// TIA Portal project "000_empty" (V21)

(* hardware
DEVICE "PLC_1"  S7-1500 station
   slot 0: "Rail_0"  Rack  6ES7 590-1***0-0AA0
   slot 1: "PLC_1"  CPU 1513-1 PN  6ES7 513-1AL02-0AB0  V2.9
      slot 3: "CPU display_1"  6ES7591-1AA00-0AA0
      slot 32768: "PROFINET interface_1"  X1
         slot 32769: "Port_1"  X1 P1
         slot 32770: "Port_2"  X1 P2
      slot 34817: "Virtual CP interface port_1"  Virtual CP interface port  Virtual CP interface port
*)

// ===== PLC "PLC_1"  CPU 1513-1 PN =====

VAR_GLOBAL   // PLC tag table "Default tag table"
   "Tag__639296449648259132" AT %MW10 : Word;
   "Tag__639296449652422717" AT %MW12 : Word;
   "Tag__639296449666761157" AT %T1 : Timer;
   "Tag__639296449667118790" AT %T2 : Timer;
   "Tag__639296449667279911" AT %T3 : Timer;
   "Tag__639296449667396582" AT %T4 : Timer;
   "Tag__639296449667490544" AT %T5 : Timer;
   "Tag__639296449667666479" AT %C1 : Counter;
END_VAR

TYPE "UDT_Motor"
   STRUCT
      Running : Bool;   // Motor on
      Speed : Real := 1500.0;   // Speed setpoint
      Count : Int := 7;
   END_STRUCT;
END_TYPE

DATA_BLOCK "DB_Global"   // DB1
{ S7_Optimized_Access := 'TRUE' }
   VAR
      xBool : Bool := TRUE;   // Bool comment
      iInt : Int := 42;
      rReal : Real := 3.5;   // Real comment
      aInt : Array[0..3] of Int;
      sData : Struct
         "a" : Bool;
         "b" : DInt := -5;
      END_STRUCT;
   END_VAR
BEGIN
   aInt[1] := 11;
END_DATA_BLOCK

DATA_BLOCK "FB_Empty_DB"   // DB2
{ S7_Optimized_Access := 'TRUE' }
VERSION : 0.1
// stored: InstanceOfName FB_Empty
"FB_Empty"
BEGIN
END_DATA_BLOCK

DATA_BLOCK "DB_Motor"   // DB4
{ S7_Optimized_Access := 'TRUE' }
   VAR
      motor : "UDT_Motor";
   END_VAR
BEGIN
   motor.Speed := 750.0;
END_DATA_BLOCK

DATA_BLOCK "FB_Iface_DB"   // DB5
{ S7_Optimized_Access := 'TRUE' }
VERSION : 0.1
// stored: InstanceOfName FB_Iface
"FB_Iface"
BEGIN
   stInt := 99;
   stBool := TRUE;
END_DATA_BLOCK

DATA_BLOCK "DB_StlStd"   // DB6
{ S7_Optimized_Access := 'FALSE' }
VERSION : 0.1
   VAR
      w0 : Word;
      w1 : Word;
   END_VAR
BEGIN
END_DATA_BLOCK

DATA_BLOCK "DB_StlInner"   // DB7
{ S7_Optimized_Access := 'TRUE' }
VERSION : 0.1
// stored: InstanceOfName FB_StlInner
"FB_StlInner"
BEGIN
END_DATA_BLOCK

// folder: BlockGroup_1

DATA_BLOCK "DB_InGroup"   // DB3
{ S7_Optimized_Access := 'TRUE' }
   VAR
      wWord : Word := 16#00FF;
   END_VAR
BEGIN
END_DATA_BLOCK

// folder: (top level)

FUNCTION_BLOCK "FB_Empty"   // FB1, SCL
{ S7_Optimized_Access := 'TRUE' }
VERSION : 0.1
BEGIN
END_FUNCTION_BLOCK

FUNCTION_BLOCK "FB_Iface"   // FB2, SCL
{ S7_Optimized_Access := 'TRUE' }
VERSION : 0.1
   VAR_INPUT
      iBool : Bool;   // Input bool
      iInt : Int;   // Input int
      iReal : Real;   // Input real
      iArr : Array[0..3] of Int;   // Input array
      iMotor : "UDT_Motor";   // Input UDT
   END_VAR
   VAR_OUTPUT
      oBool : Bool;   // Output bool
      oInt : Int;   // Output int
   END_VAR
   VAR_IN_OUT
      ioReal : Real;   // InOut real
   END_VAR
   VAR
      stInt : Int := 42;   // Static int
      stBool : Bool;   // Static bool comment
   END_VAR
   VAR_TEMP
      tInt : Int;   // Temp int
   END_VAR
   VAR CONSTANT
      cInt : Int := 7;   // Constant int
   END_VAR
BEGIN
   #tInt := #iInt + #cInt;
           #oInt := #tInt;
           #oBool := #iBool;
           #ioReal := #ioReal + #iReal;
END_FUNCTION_BLOCK

FUNCTION_BLOCK "FB_Stl"   // FB3, STL
TITLE = STL test FB
{ S7_Optimized_Access := 'TRUE' }
VERSION : 0.1
   VAR_INPUT
      start : Bool;
      stop : Bool;
   END_VAR
   VAR_OUTPUT
      running : Bool;
      count : Int;
   END_VAR
   VAR
      cnt : Int;
      edge : Bool;
   END_VAR
BEGIN

REGION Network 1: Latch
         A(;
         O     #start;
         O     #running;
         );
         AN    #stop;
         =     #running;
END_REGION

REGION Network 2: Count rising edges
         A     #start;
         FP    #edge;
         JCN   END1;
         L     #cnt;
         +     1;
         T     #cnt;
   END1: L     #cnt;
         T     #count;
         SET;
         SAVE;
END_REGION
END_FUNCTION_BLOCK

FUNCTION_BLOCK "FB_StlBe"   // FB4, STL
TITLE = STL catalog FB_StlBe
{ S7_Optimized_Access := 'TRUE' }
VERSION : 0.1
   VAR_INPUT
      "a" : Bool;
      "b" : Bool;
      c : Bool;
      i1 : Int;
      i2 : Int;
      d1 : DInt;
      d2 : DInt;
      r1 : Real;
      r2 : Real;
      w1 : Word;
      w2 : Word;
      dw1 : DWord;
      dw2 : DWord;
   END_VAR
   VAR_OUTPUT
      q : Bool;
      by1 : Byte;
      ir : Int;
      dr : DInt;
      rr : Real;
      wr : Word;
      dwr : DWord;
   END_VAR
   VAR
      dummy : Bool;
   END_VAR
BEGIN

REGION Network 1: 128 BE
         L     1;
         T     #ir;
         BE;
END_REGION
END_FUNCTION_BLOCK

FUNCTION_BLOCK "FB_StlBit"   // FB5, STL
TITLE = STL catalog FB_StlBit
{ S7_Optimized_Access := 'TRUE' }
VERSION : 0.1
   VAR_INPUT
      "a" : Bool;
      "b" : Bool;
      c : Bool;
      i1 : Int;
      i2 : Int;
      d1 : DInt;
      d2 : DInt;
      r1 : Real;
      r2 : Real;
      w1 : Word;
      w2 : Word;
      dw1 : DWord;
      dw2 : DWord;
   END_VAR
   VAR_OUTPUT
      q : Bool;
      by1 : Byte;
      ir : Int;
      dr : DInt;
      rr : Real;
      wr : Word;
      dwr : DWord;
   END_VAR
   VAR
      edgeN : Bool;
      edgeP : Bool;
   END_VAR
BEGIN

REGION Network 1: 001 A
         A     #"a";
         =     #q;
END_REGION

REGION Network 2: 002 AN
         AN    #"a";
         =     #q;
END_REGION

REGION Network 3: 003 O
         O     #"a";
         O     #"b";
         =     #q;
END_REGION

REGION Network 4: 004 ON
         ON    #"a";
         =     #q;
END_REGION

REGION Network 5: 005 X
         X     #"a";
         X     #"b";
         =     #q;
END_REGION

REGION Network 6: 006 XN
         XN    #"a";
         =     #q;
END_REGION

REGION Network 7: 007 O (2)
         A     #"a";
         A     #"b";
         O;
         A     #c;
         =     #q;
END_REGION

REGION Network 8: 008 A(
         A(;
         O     #"a";
         O     #"b";
         );
         =     #q;
END_REGION

REGION Network 9: 009 AN(
         AN(;
         O     #"a";
         O     #"b";
         );
         =     #q;
END_REGION

REGION Network 10: 010 O(
         O(;
         A     #"a";
         A     #"b";
         );
         =     #q;
END_REGION

REGION Network 11: 011 ON(
         ON(;
         A     #"a";
         );
         =     #q;
END_REGION

REGION Network 12: 012 X(
         X(;
         A     #"a";
         );
         X     #"b";
         =     #q;
END_REGION

REGION Network 13: 013 XN(
         XN(;
         A     #"a";
         );
         =     #q;
END_REGION

REGION Network 14: 014 )
         A(;
         A     #"a";
         );
         =     #q;
END_REGION

REGION Network 15: 015 =
         A     #"a";
         =     #q;
END_REGION

REGION Network 16: 016 R
         A     #"a";
         R     #q;
END_REGION

REGION Network 17: 017 S
         A     #"a";
         S     #q;
END_REGION

REGION Network 18: 018 NOT
         A     #"a";
         NOT;
         =     #q;
END_REGION

REGION Network 19: 019 SET
         SET;
         =     #q;
END_REGION

REGION Network 20: 020 CLR
         CLR;
         =     #q;
END_REGION

REGION Network 21: 021 SAVE
         A     #"a";
         SAVE;
END_REGION

REGION Network 22: 022 FN
         A     #"a";
         FN    #edgeN;
         =     #q;
END_REGION

REGION Network 23: 023 FP
         A     #"a";
         FP    #edgeP;
         =     #q;
END_REGION
END_FUNCTION_BLOCK

FUNCTION_BLOCK "FB_StlDb"   // FB6, STL
TITLE = STL catalog FB_StlDb
{ S7_Optimized_Access := 'FALSE' }
VERSION : 0.1
   VAR_INPUT
      "a" : Bool;
      "b" : Bool;
      c : Bool;
      i1 : Int;
      i2 : Int;
      d1 : DInt;
      d2 : DInt;
      r1 : Real;
      r2 : Real;
      w1 : Word;
      w2 : Word;
      dw1 : DWord;
      dw2 : DWord;
   END_VAR
   VAR_OUTPUT
      q : Bool;
      by1 : Byte;
      ir : Int;
      dr : DInt;
      rr : Real;
      wr : Word;
      dwr : DWord;
   END_VAR
   VAR
      dummy : Bool;
   END_VAR
BEGIN

REGION Network 1: 121 OPN
         OPN   "DB_StlStd";
         L     %DataW0;
         T     #wr;
         OPN   "";
END_REGION

REGION Network 2: 122 OPNDI
         OPNDI "DB_StlStd";
         L     %XDataW0;
         T     #wr;
END_REGION

REGION Network 3: 123 CDB
         CDB;
END_REGION

REGION Network 4: 124 L DBLG
         L     DBLG;
         T     #dr;
END_REGION

REGION Network 5: 125 L DBNO
         L     DBNO;
         T     #dr;
END_REGION

REGION Network 6: 126 L DILG
         L     DILG;
         T     #dr;
END_REGION

REGION Network 7: 127 L DINO
         L     DINO;
         T     #dr;
END_REGION
END_FUNCTION_BLOCK

FUNCTION_BLOCK "FB_StlInner"   // FB7, STL
{ S7_Optimized_Access := 'TRUE' }
VERSION : 0.1
   VAR_INPUT
      start : Bool;
   END_VAR
   VAR_OUTPUT
      cnt : Int;
   END_VAR
   VAR
      n : Int;
   END_VAR
BEGIN

REGION Network 1
         A     #start;
         JCN   E1;
         L     #n;
         +     1;
         T     #n;
   E1:   L     #n;
         T     #cnt;
END_REGION
END_FUNCTION_BLOCK

FUNCTION_BLOCK "FB_StlJump"   // FB8, STL
TITLE = STL catalog FB_StlJump
{ S7_Optimized_Access := 'TRUE' }
VERSION : 0.1
   VAR_INPUT
      "a" : Bool;
      "b" : Bool;
      c : Bool;
      i1 : Int;
      i2 : Int;
      d1 : DInt;
      d2 : DInt;
      r1 : Real;
      r2 : Real;
      w1 : Word;
      w2 : Word;
      dw1 : DWord;
      dw2 : DWord;
   END_VAR
   VAR_OUTPUT
      q : Bool;
      by1 : Byte;
      ir : Int;
      dr : DInt;
      rr : Real;
      wr : Word;
      dwr : DWord;
   END_VAR
   VAR
      dummy : Bool;
   END_VAR
BEGIN

REGION Network 1: 102 Jump label
         JU    LB01;
         L     1;
         T     #ir;
   LB01: NOP   0;
END_REGION

REGION Network 2: 103 JU
         JU    J001;
         L     1;
         T     #ir;
   J001: NOP   0;
END_REGION

REGION Network 3: 104 JC
         A     #"a";
         JC    J002;
         L     1;
         T     #ir;
   J002: NOP   0;
END_REGION

REGION Network 4: 105 JCN
         A     #"a";
         JCN   J003;
         L     1;
         T     #ir;
   J003: NOP   0;
END_REGION

REGION Network 5: 106 JCB
         A     #"a";
         JCB   J004;
         L     1;
         T     #ir;
   J004: NOP   0;
END_REGION

REGION Network 6: 107 JNB
         A     #"a";
         JNB   J005;
         L     1;
         T     #ir;
   J005: NOP   0;
END_REGION

REGION Network 7: 108 JBI
         A     #"a";
         SAVE;
         JBI   J006;
         L     1;
         T     #ir;
   J006: NOP   0;
END_REGION

REGION Network 8: 109 JNBI
         A     #"a";
         SAVE;
         JNBI  J007;
         L     1;
         T     #ir;
   J007: NOP   0;
END_REGION

REGION Network 9: 110 JO
         L     #i1;
         L     #i2;
         -I;
         T     #ir;
         JO    J008;
         L     1;
         T     #ir;
   J008: NOP   0;
END_REGION

REGION Network 10: 111 JOS
         L     #i1;
         L     #i2;
         -I;
         T     #ir;
         JOS   J009;
         L     1;
         T     #ir;
   J009: NOP   0;
END_REGION

REGION Network 11: 112 JZ
         L     #i1;
         L     #i2;
         -I;
         T     #ir;
         JZ    J010;
         L     1;
         T     #ir;
   J010: NOP   0;
END_REGION

REGION Network 12: 113 JN
         L     #i1;
         L     #i2;
         -I;
         T     #ir;
         JN    J011;
         L     1;
         T     #ir;
   J011: NOP   0;
END_REGION

REGION Network 13: 114 JP
         L     #i1;
         L     #i2;
         -I;
         T     #ir;
         JP    J012;
         L     1;
         T     #ir;
   J012: NOP   0;
END_REGION

REGION Network 14: 115 JM
         L     #i1;
         L     #i2;
         -I;
         T     #ir;
         JM    J013;
         L     1;
         T     #ir;
   J013: NOP   0;
END_REGION

REGION Network 15: 116 JPZ
         L     #i1;
         L     #i2;
         -I;
         T     #ir;
         JPZ   J014;
         L     1;
         T     #ir;
   J014: NOP   0;
END_REGION

REGION Network 16: 117 JMZ
         L     #i1;
         L     #i2;
         -I;
         T     #ir;
         JMZ   J015;
         L     1;
         T     #ir;
   J015: NOP   0;
END_REGION

REGION Network 17: 118 JUO
         L     #r1;
         L     #r2;
         /R;
         T     #rr;
         JUO   J016;
         L     1;
         T     #ir;
   J016: NOP   0;
END_REGION

REGION Network 18: 119 JL
         L     #i1;
         JL    LST1;
         JU    SG0;
         JU    SG1;
   LST1: JU    SEND;
   SG0:  L     10;
         T     #ir;
         JU    SEND;
   SG1:  L     11;
         T     #ir;
   SEND: NOP   0;
END_REGION

REGION Network 19: 120 LOOP
         L     5;
   NXT1: T     #ir;
         L     #ir;
         LOOP  NXT1;
END_REGION
END_FUNCTION_BLOCK

FUNCTION_BLOCK "FB_StlLoad"   // FB9, STL
TITLE = STL catalog FB_StlLoad
{ S7_Optimized_Access := 'FALSE' }
VERSION : 0.1
   VAR_INPUT
      "a" : Bool;
      "b" : Bool;
      c : Bool;
      i1 : Int;
      i2 : Int;
      d1 : DInt;
      d2 : DInt;
      r1 : Real;
      r2 : Real;
      w1 : Word;
      w2 : Word;
      dw1 : DWord;
      dw2 : DWord;
   END_VAR
   VAR_OUTPUT
      q : Bool;
      by1 : Byte;
      ir : Int;
      dr : DInt;
      rr : Real;
      wr : Word;
      dwr : DWord;
   END_VAR
   VAR
      dummy : Bool;
   END_VAR
BEGIN

REGION Network 1: 070 L
         L     #i1;
         T     #ir;
         L     "Tag__639296449648259132";
         T     #ir;
         L     P#M10.0;
         T     #dwr;
         L     B#16#12;
         T     #by1;
         L     'AB';
         T     #wr;
         L     2.5;
         T     #rr;
         L     T#1S;
         T     #dr;
END_REGION

REGION Network 2: 071 L STW
         L     STW;
         T     #wr;
END_REGION

REGION Network 3: 072 LAR1
         L     P#M10.0;
         LAR1;
END_REGION

REGION Network 4: 073 LAR1 <D>
         LAR1  P#M20.0;
         LAR1  #dw1;
END_REGION

REGION Network 5: 074 LAR1 AR2
         LAR1  AR2;
END_REGION

REGION Network 6: 075 LAR2
         L     P#M10.0;
         LAR2;
END_REGION

REGION Network 7: 076 LAR2 <D>
         LAR2  P#M30.0;
         LAR2  #dw1;
END_REGION

REGION Network 8: 077 T
         L     #i1;
         T     #ir;
         T     "Tag__639296449652422717";
         L     2;
         T     W [AR1,P#0.0];
         T     MW [#dw1];
END_REGION

REGION Network 9: 078 T STW
         L     #w1;
         T     STW;
END_REGION

REGION Network 10: 079 CAR
         CAR;
END_REGION

REGION Network 11: 080 TAR1
         TAR1;
         T     #dwr;
END_REGION

REGION Network 12: 081 TAR1 <D>
         TAR1  #dwr;
END_REGION

REGION Network 13: 082 TAR1 AR2
         TAR1  AR2;
END_REGION

REGION Network 14: 083 TAR2
         TAR2;
         T     #dwr;
END_REGION

REGION Network 15: 084 TAR2 <D>
         TAR2  #dwr;
END_REGION

REGION Network 16: 153 +AR1
         L     +4;
         +AR1;
         +AR1  P#2.0;
END_REGION

REGION Network 17: 154 +AR2
         L     +4;
         +AR2;
         +AR2  P#2.0;
END_REGION
END_FUNCTION_BLOCK

FUNCTION_BLOCK "FB_StlMath"   // FB10, STL
TITLE = STL catalog FB_StlMath
{ S7_Optimized_Access := 'TRUE' }
VERSION : 0.1
   VAR_INPUT
      "a" : Bool;
      "b" : Bool;
      c : Bool;
      i1 : Int;
      i2 : Int;
      d1 : DInt;
      d2 : DInt;
      r1 : Real;
      r2 : Real;
      w1 : Word;
      w2 : Word;
      dw1 : DWord;
      dw2 : DWord;
   END_VAR
   VAR_OUTPUT
      q : Bool;
      by1 : Byte;
      ir : Int;
      dr : DInt;
      rr : Real;
      wr : Word;
      dwr : DWord;
   END_VAR
   VAR
      dummy : Bool;
   END_VAR
BEGIN

REGION Network 1: 040 ? I
         L     #i1;
         L     #i2;
         ==I;
         =     #q;
         L     #i1;
         L     #i2;
         <>I;
         =     #q;
         L     #i1;
         L     #i2;
         >I;
         =     #q;
         L     #i1;
         L     #i2;
         <I;
         =     #q;
         L     #i1;
         L     #i2;
         >=I;
         =     #q;
         L     #i1;
         L     #i2;
         <=I;
         =     #q;
END_REGION

REGION Network 2: 041 ? D
         L     #d1;
         L     #d2;
         ==D;
         =     #q;
         L     #d1;
         L     #d2;
         <>D;
         =     #q;
         L     #d1;
         L     #d2;
         >D;
         =     #q;
         L     #d1;
         L     #d2;
         <D;
         =     #q;
         L     #d1;
         L     #d2;
         >=D;
         =     #q;
         L     #d1;
         L     #d2;
         <=D;
         =     #q;
END_REGION

REGION Network 3: 042 ? R
         L     #r1;
         L     #r2;
         ==R;
         =     #q;
         L     #r1;
         L     #r2;
         <>R;
         =     #q;
         L     #r1;
         L     #r2;
         >R;
         =     #q;
         L     #r1;
         L     #r2;
         <R;
         =     #q;
         L     #r1;
         L     #r2;
         >=R;
         =     #q;
         L     #r1;
         L     #r2;
         <=R;
         =     #q;
END_REGION

REGION Network 4: 043 +I
         L     #i1;
         L     #i2;
         +I;
         T     #ir;
END_REGION

REGION Network 5: 044 -I
         L     #i1;
         L     #i2;
         -I;
         T     #ir;
END_REGION

REGION Network 6: 045 *I
         L     #i1;
         L     #i2;
         *I;
         T     #ir;
END_REGION

REGION Network 7: 046 /I
         L     #i1;
         L     #i2;
         /I;
         T     #ir;
END_REGION

REGION Network 8: 047 +D
         L     #d1;
         L     #d2;
         +D;
         T     #dr;
END_REGION

REGION Network 9: 048 -D
         L     #d1;
         L     #d2;
         -D;
         T     #dr;
END_REGION

REGION Network 10: 049 *D
         L     #d1;
         L     #d2;
         *D;
         T     #dr;
END_REGION

REGION Network 11: 050 /D
         L     #d1;
         L     #d2;
         /D;
         T     #dr;
END_REGION

REGION Network 12: 051 +
         L     #i1;
         +     5;
         T     #ir;
END_REGION

REGION Network 13: 052 INC
         L     #by1;
         INC   1;
         T     #by1;
END_REGION

REGION Network 14: 053 DEC
         L     #by1;
         DEC   1;
         T     #by1;
END_REGION

REGION Network 15: 054 MOD
         L     #d1;
         L     #d2;
         MOD;
         T     #dr;
END_REGION

REGION Network 16: 055 +R
         L     #r1;
         L     #r2;
         +R;
         T     #rr;
END_REGION

REGION Network 17: 056 -R
         L     #r1;
         L     #r2;
         -R;
         T     #rr;
END_REGION

REGION Network 18: 057 *R
         L     #r1;
         L     #r2;
         *R;
         T     #rr;
END_REGION

REGION Network 19: 058 /R
         L     #r1;
         L     #r2;
         /R;
         T     #rr;
END_REGION

REGION Network 20: 059 ABS
         L     #r1;
         ABS;
         T     #rr;
END_REGION

REGION Network 21: 060 SQR
         L     #r1;
         SQR;
         T     #rr;
END_REGION

REGION Network 22: 061 SQRT
         L     #r1;
         SQRT;
         T     #rr;
END_REGION

REGION Network 23: 062 EXP
         L     #r1;
         EXP;
         T     #rr;
END_REGION

REGION Network 24: 063 LN
         L     #r1;
         LN;
         T     #rr;
END_REGION

REGION Network 25: 064 SIN
         L     #r1;
         SIN;
         T     #rr;
END_REGION

REGION Network 26: 065 ASIN
         L     #r1;
         ASIN;
         T     #rr;
END_REGION

REGION Network 27: 066 COS
         L     #r1;
         COS;
         T     #rr;
END_REGION

REGION Network 28: 067 ACOS
         L     #r1;
         ACOS;
         T     #rr;
END_REGION

REGION Network 29: 068 TAN
         L     #r1;
         TAN;
         T     #rr;
END_REGION

REGION Network 30: 069 ATAN
         L     #r1;
         ATAN;
         T     #rr;
END_REGION

REGION Network 31: 085 BTI
         L     #w1;
         BTI;
         T     #ir;
END_REGION

REGION Network 32: 086 ITB
         L     #i1;
         ITB;
         T     #wr;
END_REGION

REGION Network 33: 087 BTD
         L     #dw1;
         BTD;
         T     #dr;
END_REGION

REGION Network 34: 088 ITD
         L     #i1;
         ITD;
         T     #dr;
END_REGION

REGION Network 35: 089 DTB
         L     #d1;
         DTB;
         T     #dwr;
END_REGION

REGION Network 36: 090 DTR
         L     #d1;
         DTR;
         T     #rr;
END_REGION

REGION Network 37: 091 INVI
         L     #i1;
         INVI;
         T     #ir;
END_REGION

REGION Network 38: 092 INVD
         L     #d1;
         INVD;
         T     #dr;
END_REGION

REGION Network 39: 093 NEGI
         L     #i1;
         NEGI;
         T     #ir;
END_REGION

REGION Network 40: 094 NEGD
         L     #d1;
         NEGD;
         T     #dr;
END_REGION

REGION Network 41: 095 NEGR
         L     #r1;
         NEGR;
         T     #rr;
END_REGION

REGION Network 42: 096 CAW
         L     #w1;
         CAW;
         T     #wr;
END_REGION

REGION Network 43: 097 CAD
         L     #dw1;
         CAD;
         T     #dwr;
END_REGION

REGION Network 44: 098 RND
         L     #r1;
         RND;
         T     #dr;
END_REGION

REGION Network 45: 099 TRUNC
         L     #r1;
         TRUNC;
         T     #dr;
END_REGION

REGION Network 46: 100 RND+
         L     #r1;
         RND+;
         T     #dr;
END_REGION

REGION Network 47: 101 RND-
         L     #r1;
         RND-;
         T     #dr;
END_REGION

REGION Network 48: 134 AW
         L     #w1;
         L     #w2;
         AW;
         T     #wr;
         L     #w1;
         AW    W#16#00FF;
         T     #wr;
END_REGION

REGION Network 49: 135 OW
         L     #w1;
         L     #w2;
         OW;
         T     #wr;
         L     #w1;
         OW    W#16#00FF;
         T     #wr;
END_REGION

REGION Network 50: 136 XOW
         L     #w1;
         L     #w2;
         XOW;
         T     #wr;
         L     #w1;
         XOW   W#16#00FF;
         T     #wr;
END_REGION

REGION Network 51: 137 AD
         L     #dw1;
         L     #dw2;
         AD;
         T     #dwr;
         L     #dw1;
         AD    DW#16#0000_FFFF;
         T     #dwr;
END_REGION

REGION Network 52: 138 OD
         L     #dw1;
         L     #dw2;
         OD;
         T     #dwr;
         L     #dw1;
         OD    DW#16#0000_FFFF;
         T     #dwr;
END_REGION

REGION Network 53: 139 XOD
         L     #dw1;
         L     #dw2;
         XOD;
         T     #dwr;
         L     #dw1;
         XOD   DW#16#0000_FFFF;
         T     #dwr;
END_REGION

REGION Network 54: 140 SSI
         L     #i1;
         SSI   2;
         T     #ir;
         L     2;
         L     #i1;
         SSI;
         T     #ir;
END_REGION

REGION Network 55: 141 SSD
         L     #d1;
         SSD   2;
         T     #dr;
         L     2;
         L     #d1;
         SSD;
         T     #dr;
END_REGION

REGION Network 56: 142 SLW
         L     #w1;
         SLW   2;
         T     #wr;
         L     2;
         L     #w1;
         SLW;
         T     #wr;
END_REGION

REGION Network 57: 143 SRW
         L     #w1;
         SRW   2;
         T     #wr;
         L     2;
         L     #w1;
         SRW;
         T     #wr;
END_REGION

REGION Network 58: 144 SLD
         L     #dw1;
         SLD   2;
         T     #dwr;
         L     2;
         L     #dw1;
         SLD;
         T     #dwr;
END_REGION

REGION Network 59: 145 SRD
         L     #dw1;
         SRD   2;
         T     #dwr;
         L     2;
         L     #dw1;
         SRD;
         T     #dwr;
END_REGION

REGION Network 60: 146 RLD
         L     #dw1;
         RLD   3;
         T     #dwr;
END_REGION

REGION Network 61: 147 RRD
         L     #dw1;
         RRD   3;
         T     #dwr;
END_REGION

REGION Network 62: 148 RLDA
         L     #dw1;
         RLDA;
         T     #dwr;
END_REGION

REGION Network 63: 149 RRDA
         L     #dw1;
         RRDA;
         T     #dwr;
END_REGION

REGION Network 64: 150 TAK
         L     #i1;
         L     #i2;
         TAK;
         T     #ir;
END_REGION

REGION Network 65: 151 PUSH
         L     #i1;
         PUSH;
         T     #ir;
END_REGION

REGION Network 66: 152 POP
         L     #i1;
         L     #i2;
         POP;
         T     #ir;
END_REGION

REGION Network 67: 155 BLD
         BLD   100;
END_REGION

REGION Network 68: 156 NOP 0
         NOP   0;
END_REGION

REGION Network 69: 157 NOP 1
         NOP   1;
END_REGION
END_FUNCTION_BLOCK

FUNCTION_BLOCK "FB_StlTimer"   // FB11, STL
TITLE = STL catalog FB_StlTimer
{ S7_Optimized_Access := 'TRUE' }
VERSION : 0.1
   VAR_INPUT
      "a" : Bool;
      "b" : Bool;
      c : Bool;
      i1 : Int;
      i2 : Int;
      d1 : DInt;
      d2 : DInt;
      r1 : Real;
      r2 : Real;
      w1 : Word;
      w2 : Word;
      dw1 : DWord;
      dw2 : DWord;
   END_VAR
   VAR_OUTPUT
      q : Bool;
      by1 : Byte;
      ir : Int;
      dr : DInt;
      rr : Real;
      wr : Word;
      dwr : DWord;
   END_VAR
   VAR
      dummy : Bool;
   END_VAR
BEGIN

REGION Network 1: 024 FR
         A     #"a";
         FR    "Tag__639296449666761157";
END_REGION

REGION Network 2: 025 L
         L     "Tag__639296449666761157";
         T     #wr;
END_REGION

REGION Network 3: 026 LC
         LC    "Tag__639296449666761157";
         T     #wr;
END_REGION

REGION Network 4: 027 R
         A     #"a";
         R     "Tag__639296449666761157";
END_REGION

REGION Network 5: 028 SP
         A     #"a";
         L     S5T#1S;
         SP    "Tag__639296449666761157";
END_REGION

REGION Network 6: 029 SE
         A     #"a";
         L     S5T#2S;
         SE    "Tag__639296449667118790";
END_REGION

REGION Network 7: 030 SD
         A     #"a";
         L     S5T#3S;
         SD    "Tag__639296449667279911";
END_REGION

REGION Network 8: 031 SS
         A     #"a";
         L     S5T#4S;
         SS    "Tag__639296449667396582";
END_REGION

REGION Network 9: 032 SF
         A     #"a";
         L     S5T#5S;
         SF    "Tag__639296449667490544";
END_REGION

REGION Network 10: 033 FR
         A     #"a";
         FR    "Tag__639296449667666479";
END_REGION

REGION Network 11: 034 L
         L     "Tag__639296449667666479";
         T     #wr;
END_REGION

REGION Network 12: 035 LC
         LC    "Tag__639296449667666479";
         T     #wr;
END_REGION

REGION Network 13: 036 R
         A     #"a";
         R     "Tag__639296449667666479";
END_REGION

REGION Network 14: 037 S
         A     #"a";
         L     C#5;
         S     "Tag__639296449667666479";
END_REGION

REGION Network 15: 038 CU
         A     #"a";
         CU    "Tag__639296449667666479";
END_REGION

REGION Network 16: 039 CD
         A     #"a";
         CD    "Tag__639296449667666479";
END_REGION
END_FUNCTION_BLOCK

FUNCTION_BLOCK "FB_StlCall"   // FB12, STL
TITLE = STL catalog FB_StlCall
{ S7_Optimized_Access := 'TRUE' }
VERSION : 0.1
   VAR_INPUT
      "a" : Bool;
      "b" : Bool;
      c : Bool;
      i1 : Int;
      i2 : Int;
      d1 : DInt;
      d2 : DInt;
      r1 : Real;
      r2 : Real;
      w1 : Word;
      w2 : Word;
      dw1 : DWord;
      dw2 : DWord;
   END_VAR
   VAR_OUTPUT
      q : Bool;
      by1 : Byte;
      ir : Int;
      dr : DInt;
      rr : Real;
      wr : Word;
      dwr : DWord;
   END_VAR
   VAR
      inner : "FB_StlInner";
   END_VAR
BEGIN

REGION Network 1: 129 BEC
         A     #"a";
         BEC;
END_REGION

REGION Network 2: 130 BEU
         A     #"b";
         JCN   NBEU;
         BEU;
   NBEU: NOP   0;
END_REGION

REGION Network 3: 131 CALL
         CALL  "FC_StlPar"
         ( x := #i1,
           y := 5,
           q := #q,
           r := #ir
         );
         CALL  #inner
         ( start := #"a",
           cnt   := #ir
         );
         CALL  "FB_StlInner", "DB_StlInner"
         ( start := #"b",
           cnt   := #ir
         );
END_REGION

REGION Network 4: 132 CC
         A     #"a";
         CC    "FC_StlNoPar";
END_REGION

REGION Network 5: 133 UC
         UC    "FC_StlNoPar";
END_REGION
END_FUNCTION_BLOCK

FUNCTION "FC_Stl" : Void   // FC1, STL
TITLE = STL test FC
{ S7_Optimized_Access := 'TRUE' }
VERSION : 0.1
   VAR_INPUT
      "a" : Bool;
      "b" : Bool;
      x : Int;
      y : Int;
   END_VAR
   VAR_OUTPUT
      q : Bool;
      sum : Int;
   END_VAR
   VAR_TEMP
      t : Int;
   END_VAR
BEGIN

REGION Network 1: Bit logic
   // Network comment line 1
         A     #"a";  // and a
         AN    #"b";
         =     #q;
END_REGION

REGION Network 2: Arithmetic
         L     #x;
         L     #y;
         +I;
         T     #t;

         L     #t;
         L     0;
         >I;
         JC    M001;
         L     0;
         T     #t;
   M001: L     #t;
         T     #sum;
END_REGION
END_FUNCTION

FUNCTION "FC_StlNoPar" : Void   // FC2, STL
{ S7_Optimized_Access := 'FALSE' }
VERSION : 0.1
BEGIN

REGION Network 1
         NOP   0;
END_REGION
END_FUNCTION

FUNCTION "FC_StlPar" : Void   // FC3, STL
{ S7_Optimized_Access := 'TRUE' }
VERSION : 0.1
   VAR_INPUT
      x : Int;
      y : Int;
   END_VAR
   VAR_OUTPUT
      q : Bool;
      r : Int;
   END_VAR
BEGIN

REGION Network 1
         L     #x;
         L     #y;
         +I;
         T     #r;
         >I;
         =     #q;
END_REGION
END_FUNCTION

ORGANIZATION_BLOCK "Main"   // OB1, LAD, ProgramCycle
TITLE = "Main Program Sweep (Cycle)"
{ S7_Optimized_Access := 'TRUE' }
VERSION : 0.1
   VAR_INPUT
      Initial_Call : Bool;   // Initial call of this OB
      Remanence : Bool;   // =True, if remanent data are available
   END_VAR
BEGIN
END_ORGANIZATION_BLOCK